(* Logix 5000 project; controller DSFW_0512_C_FCB_S1_SPN vendor 1 type 14 code 77 rev 20.12; software revision 20.06 *)

TASK MainTask (continuous, watchdog 500 ms) : General_Alarms_Config, Process_Control
TASK PID_Loops (periodic, rate 10 ms, priority 10, watchdog 500 ms) : Process_PID_Calculations

MODULES
   Controller : vendor 1 type 14 code 77 (CompactLogixL32EController 0, rev 20.12)
      LocalENB : 1769-L32E Ethernet Port (CompactLogixL32Ethernet 1, Ethernet 192.168.1.30, rev 20.11)
      Local : CompactBus (CompactVirtualAdapter 3, rev 20.11)
          : vendor 1 type 7 code 82 (Compact 1, rev 1.1, Input RPI 20 ms)
          : 1769-IF8 (Compact 3, rev 1.1, Output RPI 80 ms)
          : 1769-IR6 (Compact 4, rev 1.1, Input RPI 5 ms)
          : vendor 1 type 7 code 93 (Compact 2, rev 1.1, Output RPI 20 ms)
          : vendor 1 type 10 code 39 (Compact 5, rev 2.1, Output RPI 80 ms)
END_MODULES

VAR_GLOBAL   (* controller tags *)
   Alarms : DINT[3] := ([0] := 2);
   Alarms_Active : BOOL := 1;
   Batch_Mode_Enable : BOOL;
   Comp_Low_Pressure_Alarm_Setpoint : REAL := 12.0;
   Compressor_High_Pressure_Alarm_Setpoint : REAL := 300.0;
   Compressor_High_Pressure_Delay_Timer : TIMER := (PRE := 1000);
   Compressor_High_Superheat_Alarm_Delay : TIMER := (PRE := 600000);
   Compressor_High_Superheat_Alarm_Setpoint : REAL := 80.0;
   Compressor_Low_Pressure_Alarm_Setpoint : DINT := 120;
   Compressor_Low_Pressure_Delay_Timer : TIMER := (PRE := 60000);
   Compressor_Low_Subcooling_Alarm_Delay : TIMER := (PRE := 600000);
   Compressor_Low_Subcooling_Alarm_Setpoint : REAL := 4.0;
   Compressor_Low_Superheat_Alarm_Delay : TIMER := (PRE := 120000);
   Compressor_Low_Superheat_Alarm_Setpoint : REAL := 2.0;
   Compressor_OK_To_Run : BOOL;
   Compressor_Run_Proof_Delay : TIMER := (PRE := 5000);
   Compressor_Short_Cycle_Time_Remaining : REAL;
   Compressor_Short_Cycle_Timer : TIMER := (PRE := 60000);
   Compressor_Start_Delay : TIMER := (PRE := 10000);
   Compressor_Subcooling : REAL := 7.55085;
   Compressor_Superheat : REAL := 32.681896;
   Compresssor_Status : BOOL;
   Critical_Alarm : BOOL;
   DeltaV_Online : BOOL := 1;
   DeltaV_Status : DINT := 3;
   Display_Vessel_Select : BOOL;
   DV_IN_F8_50_99 : REAL[10] := ([0] := 11.0, [1] := 21.0, [2] := 21.0, [3] := 21.0); {produced}
   DV_IN_N7_100_199 : INT[10] := ([0] := 20, [1] := 4); {produced}
   DV_OUT_F8_0_49 : REAL[20] := ([0] := 21.3, [1] := 21.2, [2] := 10.7202635, [3] := -37.5, [4] := -37.5, [5] := -37.5, [8] := 109.89375, [9] := 180.79688, [10] := 79.402695, [11] := 8.548732, [13] := 74.6, [14] := 73.2, [15] := 84.7); {produced, access Read Only}
   DV_OUT_N7_0_99 : INT[20] := ([0] := 41, [1] := 16845, [2] := 3, [3] := 1, [4] := 2); {produced, access Read Only}
   EEV_101_Auto_Manual : BOOL;
   EEV_101_Manual_Output : REAL := 25.0;
   EEV_101_Output_Percent : REAL;
   EEV_101_Pressure_PIDE : PID_ENHANCED := (PV := 10.73405, PVEUMax := 103.0, PVEUMin := -7.3, SPProg := 125.0, SPOper := 125.0, SPHLimit := 103.0, SPLLimit := -7.3, RatioProg := 1.0, RatioOper := 1.0, RatioHLimit := 1.0, RatioLLimit := 1.0, CVEUMax := 10000.0, CVHLimit := 100.0, CVLLimit := 20.0, HandFB := 25.0, PGain := 10.0, IGain := 5.0, PVEDerivative := 1, ProgOverrideReq := 1, RTSTime := 1, CVLAlarm := 1, SP := 103.0, SPPercent := 100.0, SPHAlarm := 1, PVPercent := 16.35, E := 92.26595, EPercent := 83.65, InitPrimary := 1, WindupHOut := 1, WindupLOut := 1, Ratio := 1.0, Override := 1, DeltaT := 0.01, Status1 := 16#0000_0061, InstructFault := 1, SPProgInv := 1, SPOperInv := 1);
   EEV_101_Pressure_Setpoint : REAL := 125.0;
   EEV_101_Range_1_Max : REAL := 100.0;
   EEV_101_Range_1_Min : REAL := 20.0;
   EEV_101_Range_2_Max : REAL := 100.0;
   EEV_101_Range_2_Min : REAL := 20.0;
   EEV_101_Range_3_Max : REAL := 50.0;
   EEV_101_Range_3_Min : REAL := 10.0;
   EEV_101_Run_PIDE : BOOL;
   EEV_101_Run_Temp_PIDE : BOOL;
   EEV_101_Stop_PIDE : BOOL := 1;
   EEV_101_Superheat_PIDE : PID_ENHANCED := (PV := 21.081898, PVEUMax := 121.0, PVEUMin := -18.0, SPProg := 10.0, SPOper := 10.0, SPHLimit := 121.0, SPLLimit := -18.0, RatioProg := 1.0, RatioOper := 1.0, RatioHLimit := 1.0, RatioLLimit := 1.0, CVEUMax := 10000.0, CVHLimit := 100.0, CVLLimit := 20.0, HandFB := 25.0, ControlAction := 1, PGain := 10.0, IGain := 5.0, PVEDerivative := 1, ProgOverrideReq := 1, RTSTime := 1, CVLAlarm := 1, SP := 10.0, SPPercent := 20.143885, PVPercent := 28.116474, E := 11.081898, EPercent := 7.9725895, InitPrimary := 1, WindupHOut := 1, Ratio := 1.0, Override := 1, DeltaT := 0.01);
   EEV_101_Superheat_Setpoint : REAL := 10.0;
   EEV_101_Temperature_PIDE : PID_ENHANCED := (PV := 21.3, PVEUMax := 121.0, PVEUMin := -18.0, SPProg := 11.0, SPOper := 11.0, SPCascade := 11.0, SPHLimit := 121.0, SPLLimit := -18.0, RatioProg := 1.0, RatioOper := 1.0, RatioHLimit := 1.0, RatioLLimit := 1.0, CVEUMax := 10000.0, CVHLimit := 100.0, CVLLimit := 20.0, HandFB := 25.0, ControlAction := 1, PGain := 10.0, IGain := 5.0, PVEDerivative := 1, AllowCasRat := 1, ProgOverrideReq := 1, RTSTime := 1, CVLAlarm := 1, SP := 11.0, SPPercent := 20.86331, PVPercent := 28.27338, E := 10.299999, EPercent := 7.4100704, InitPrimary := 1, WindupHOut := 1, Ratio := 1.0, Override := 1, DeltaT := 0.01);
   EEV_102_Auto_Manual : BOOL;
   EEV_102_Manual_Output : REAL := 12.0;
   EEV_102_Output_Percent : REAL;
   EEV_102_PIDE : PID_ENHANCED := (PV := 32.681896, PVEUMax := 121.0, PVEUMin := -18.0, SPProg := 50.0, SPOper := 50.0, SPHLimit := 121.0, SPLLimit := -18.0, RatioProg := 1.0, RatioOper := 1.0, RatioHLimit := 1.0, RatioLLimit := 1.0, CVEUMax := 10000.0, CVHLimit := 100.0, HandFB := 12.0, ControlAction := 1, PGain := 0.3, IGain := 0.1, PVEDerivative := 1, ProgOverrideReq := 1, RTSTime := 1, SP := 50.0, SPPercent := 48.920864, PVPercent := 36.461796, E := -17.318104, EPercent := -12.459068, InitPrimary := 1, Ratio := 1.0, Override := 1, DeltaT := 0.01);
   EEV_102_SH_Setpoint : REAL := 50.0;
   EEV_102_Stop_PIDE : BOOL := 1;
   Enable_Batch : BOOL := 1;
   Evaporator_Low_Flow_Delay_Timer : TIMER;
   Evaporator_Low_Flow_Setpoint : REAL;
   Evaporator_Low_Superheat_Alarm_Delay : TIMER := (PRE := 120);
   Evaporator_Low_Superheat_Alarm_Setpoint : REAL;
   Evaporator_Superheat : REAL := 21.081898;
   Glycol_Skid_Run : BOOL;
   Glycol_Skid_Status : BOOL;
   Heater_Start_Delay : TIMER := (PRE := 5000);
   Heaters_OK_To_Run : BOOL;
   HMI_Compressor_High_Superheat_Delay : REAL := 600.0;
   HMI_Compressor_Low_Pressure_Delay : REAL := 60.0;
   HMI_Compressor_Low_Subcooling_Delay : REAL := 600.0;
   HMI_Compressor_Low_Superheat_Delay : REAL := 120.0;
   HMI_Evaporator_Low_Superheat_Delay : REAL := 120.0;
   HMI_Pump_High_Pressure_Delay : REAL;
   HMI_Pump_Low_Pressure_Delay : REAL := 20.0;
   HMI_Remote_Enable : BOOL := 1;
   HMI_Tank_High_Pressure_Delay : REAL := 5.0;
   HMI_Tank_Low_Level_Delay : REAL := 10.0;
   Jacket_High_High_Temperature_Setpoint : REAL := 110.0;
   Jacket_High_Temperature_Setpoint : REAL := 110.0;
   Jacket_Low_Low_Temperature_Setpoint : REAL := -20.0;
   Jacket_Low_Temperature_Setpoint : REAL := -20.0;
   Large_Batch_Derivative : REAL;
   Large_Batch_Integral : REAL := 0.9;
   Large_Batch_Proportional : REAL := 15.0;
   Large_Batch_Selected : BOOL;
   LSH_101_Status : BOOL := 1;
   LSL_101_Status : BOOL := 1;
   LSL_102_Status : BOOL := 1;
   Medium_Batch_Derivative : REAL;
   Medium_Batch_Integral : REAL := 0.9;
   Medium_Batch_Proportional : REAL := 15.0;
   Medium_Batch_Selected : BOOL;
   Phase_Monitor_Delay : TIMER := (PRE := 5000);
   Process_Pump_Flow_Rate : REAL := -45.73986;
   Process_Pump_Low_Flow_Alarm_Setpoint : DINT;
   PT_101_Offset : REAL;
   PT_101_Reactor_Supply_Pressure : REAL := 10.713368;
   PT_101_Sensor_Alarm_Delay : TIMER := (PRE := 5000);
   PT_102_Compressor_Suction_Pressure : REAL := 109.89375;
   PT_102_Offset : REAL;
   PT_102_Sensor_Alarm_Delay : TIMER := (PRE := 5000);
   PT_103_Compressor_Discharge_Pressure : REAL := 180.79688;
   PT_103_Offset : REAL;
   PT_103_Sensor_Alarm_Delay : TIMER := (PRE := 5000);
   PT_104_Evaporator_Suction_Pressure : REAL := 109.89375;
   PT_104_Offset : REAL;
   PT_104_Sensor_Alarm_Delay : TIMER := (PRE := 5000);
   PT_105_Offset : REAL;
   PT_105_Sensor_Alarm_Delay : TIMER := (PRE := 5000);
   PT_105_Tank_Blanket_Pressure : REAL := 8.562519;
   Pump_High_Pressure_Delay : TIMER;
   Pump_High_Pressure_Setpoint : REAL := 100.0;
   Pump_Low_Flow_Delay_Timer : TIMER;
   Pump_Low_Pressure_Delay : TIMER := (PRE := 20000);
   Pump_Low_Pressure_Setpoint : REAL := 5.0;
   Pump_OK_To_Run : BOOL;
   Pump_Start_Delay : TIMER := (PRE := 5000);
   Pump_Status : BOOL;
   Reaactor_Batch_PIDE : PID_ENHANCED := (PV := -37.5, PVEUMax := 100.0, PVEUMin := -15.0, SPProg := 11.0, SPOper := -15.0, SPHLimit := 100.0, SPLLimit := -15.0, RatioProg := 1.0, RatioOper := 1.0, RatioHLimit := 1.0, RatioLLimit := 1.0, CVInitReq := 1, CVInitValue := 11.0, CVEUMax := -32.5, CVEUMin := -5.0, CVHLimit := 100.0, PGain := 15.0, IGain := 0.9, PVEDerivative := 1, DSmoothing := 1, PVTracking := 1, ManualAfterInit := 1, ProgOverrideReq := 1, RTSTime := 1, CVEU := 11.0, CVInitializing := 1, CVLAlarm := 1, SP := -15.0, SPLAlarm := 1, PVPercent := -19.565218, E := 22.5, EPercent := 19.565218, InitPrimary := 1, Ratio := 1.0, Override := 1, DeltaT := 0.01);
   Reactor_Batch_CV_as_SP : REAL := 11.0;
   Reactor_Batch_PID_Start : BOOL;
   Reactor_Batch_PID_Start_Delay : TIMER := (PRE := 5000);
   Reactor_Batch_PID_Start_ONS : BOOL;
   Reactor_Batch_PID_Stop : BOOL := 1;
   Reactor_Batch_PV : REAL := -37.5;
   Reactor_Batch_SP_High : REAL := -32.5;
   Reactor_Batch_SP_Low : REAL := -42.5;
   Read_PLC_Clock : DINT[7] := ([0] := 1999, [1] := 12, [2] := 29, [3] := 18, [4] := 28, [5] := 41, [6] := 799818);
   Remote_Enable : BOOL := 1;
   Remote_Start : BOOL;
   Reset_Alarms : BOOL;
   Reset_Defaults : BOOL;
   SCR_101_Auto_Manual : BOOL;
   SCR_101_Manual_Output : REAL;
   SCR_101_Output_Percent : REAL;
   SCR_101_PIDE : PID_ENHANCED := (PV := 21.3, PVEUMax := 121.0, PVEUMin := -18.0, SPProg := 11.0, SPOper := 21.3, SPCascade := 11.0, SPHLimit := 121.0, SPLLimit := -18.0, RatioProg := 1.0, RatioOper := 1.0, RatioHLimit := 1.0, RatioLLimit := 1.0, CVEUMax := 10000.0, CVHLimit := 100.0, PGain := 50.0, IGain := 5.0, PVEDerivative := 1, PVTracking := 1, AllowCasRat := 1, ProgOverrideReq := 1, RTSTime := 1, SP := 21.3, SPPercent := 28.27338, PVPercent := 28.27338, InitPrimary := 1, Ratio := 1.0, Override := 1, DeltaT := 0.01);
   SCR_101_Run_PIDE : BOOL;
   SCR_101_Stop_PIDE : BOOL := 1;
   Select_Large_Batch : BOOL;
   Select_Medium_Batch : BOOL;
   Select_Small_Batch : BOOL;
   Select_Vessel_1 : BOOL;
   Select_Vessel_2 : BOOL;
   Select_Vessel_3 : BOOL;
   Show_Local : BOOL;
   SIC_101_Auto_Manual : BOOL;
   SIC_101_Manual_Output : REAL := 100.0;
   SIC_101_Output_Percent : REAL;
   SIC_101_PIDE : PID_ENHANCED := (PV := 10.740945, PVEUMax := 103.0, PVEUMin := -7.3, SPProg := 50.0, SPOper := 50.0, SPHLimit := 103.0, SPLLimit := -7.3, RatioProg := 1.0, RatioOper := 1.0, RatioHLimit := 1.0, RatioLLimit := 1.0, CVEUMax := 10000.0, CVHLimit := 100.0, HandFB := 100.0, IGain := 10.0, PVEDerivative := 1, ProgOverrideReq := 1, RTSTime := 1, SP := 50.0, SPPercent := 51.949226, PVPercent := 16.35625, E := 39.259056, EPercent := 35.592976, InitPrimary := 1, Ratio := 1.0, Override := 1, DeltaT := 0.01);
   SIC_101_Pressure_Setpoint : REAL := 50.0;
   SIC_101_Run_PIDE : BOOL;
   SIC_101_Stop_PIDE : BOOL := 1;
   Small_Batch_Derivative : REAL;
   Small_Batch_Integral : REAL := 0.9;
   Small_Batch_Proportional : REAL := 15.0;
   Small_Batch_Selected : BOOL;
   SP_Add_Max : REAL := 5.0;
   SP_Add_Min : REAL := 50.0;
   Startup_Delay : TIMER := (PRE := 250, ACC := 250, EN := 1, DN := 1);
   System_Start : BOOL := 1;
   Tank_High_Pressure_Delay : TIMER := (PRE := 5000);
   Tank_High_Pressure_Setpoint : REAL := 15.0;
   Tank_Low_Level_Delay : TIMER := (PRE := 10000);
   TCV_101_Auto_Manual : BOOL;
   TCV_101_Define_Range_1_Max : REAL := -5.0;
   TCV_101_Define_Range_1_Min : REAL := -30.0;
   TCV_101_Define_Range_2_Max : REAL := 50.0;
   TCV_101_Define_Range_2_Min : REAL := -4.9;
   TCV_101_Define_Range_3_Max : REAL := 130.0;
   TCV_101_Define_Range_3_Min : REAL := 50.1;
   TCV_101_Manual_Output : REAL;
   TCV_101_Output_Percent : REAL;
   TCV_101_PIDE : PID_ENHANCED := (PV := 21.3, PVEUMax := 121.0, PVEUMin := -18.0, SPProg := 11.0, SPOper := 11.0, SPCascade := 11.0, SPHLimit := 121.0, SPLLimit := -18.0, RatioProg := 1.0, RatioOper := 1.0, RatioHLimit := 1.0, RatioLLimit := 1.0, CVEUMax := 10000.0, CVHLimit := 50.0, CVLLimit := 15.0, PGain := 10.0, IGain := 5.0, PVEDerivative := 1, AllowCasRat := 1, ProgOverrideReq := 1, RTSTime := 1, CVLAlarm := 1, SP := 11.0, SPPercent := 20.86331, PVPercent := 28.27338, E := -10.299999, EPercent := -7.4100704, InitPrimary := 1, WindupLOut := 1, Ratio := 1.0, Override := 1, DeltaT := 0.01);
   TCV_101_Range_1_Max : REAL := 50.0;
   TCV_101_Range_1_Min : REAL := 15.0;
   TCV_101_Range_2_Max : REAL := 50.0;
   TCV_101_Range_2_Min : REAL := 15.0;
   TCV_101_Range_3_Max : REAL := 50.0;
   TCV_101_Range_3_Min : REAL := 5.0;
   TCV_101_Run_PIDE : BOOL;
   TCV_101_Stop_PIDE : BOOL := 1;
   TE_101_Liquid_Line_Temperature : REAL := 74.6;
   TE_101_Offset : REAL;
   TE_102_Evaporator_Suction_Temperature : REAL := 73.1;
   TE_102_Offset : REAL;
   TE_103_Compressor_Suction_Temperature : REAL := 84.6;
   TE_103_Offset : REAL;
   TE_104_Offset : REAL;
   TE_104_Reactor_Return_Temperature : REAL := 21.2;
   TE_105_Offset : REAL;
   TE_105_Reactor_Supply_Temperature : REAL := 21.3;
   Temperature_Setpoint : REAL := 11.0;
   Test_Analog : REAL := 4000.0;
   Test_Bit : BOOL[32] := ([0] := 1, [1] := 1);
   TIT_101_Offset : REAL;
   TIT_101_Sensor_Alarm_Delay : TIMER := (PRE := 5000);
   TIT_101_Vessel_Temperature : REAL := -37.5;
   TIT_201_Offset : REAL;
   TIT_201_Sensor_Alarm_Delay : TIMER;
   TIT_201_Vessel_Temperature : REAL := -37.5;
   TIT_301_Offset : REAL;
   TIT_301_Sensor_Alarm_Delay : TIMER;
   TIT_301_Vessel_Temperature : REAL := -37.5;
   Vessel_1_Scale_Max : REAL := 120.0;
   Vessel_1_Scale_Min : REAL := -30.0;
   Vessel_1_Selected : BOOL;
   Vessel_2_Scale_Max : REAL := 120.0;
   Vessel_2_Scale_Min : REAL := -30.0;
   Vessel_2_Selected : BOOL;
   Vessel_3_Scale_Max : REAL := 120.0;
   Vessel_3_Scale_Min : REAL := -30.0;
   Vessel_3_Selected : BOOL;
   Vessel_High_High_Temperature_Setpoint : REAL := 110.0;
   Vessel_High_Temperature_Setpoint : REAL := 110.0;
   Vessel_Low_Low_Temperature_Setpoint : REAL := -20.0;
   Vessel_Low_Temperature_Setpoint : REAL := -20.0;
   Warning_Alarms : BOOL := 1;
END_VAR

PROGRAM General_Alarms_Config   (* main routine MainRoutine *)

ROUTINE DV_Communications   (* ladder *)
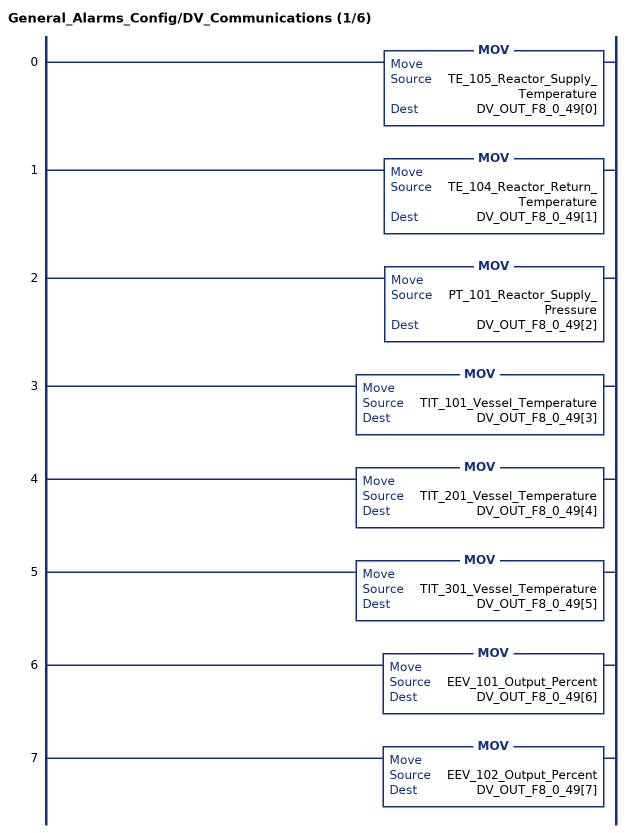
   0: MOV(TE_105_Reactor_Supply_Temperature,DV_OUT_F8_0_49[0]);
   1: MOV(TE_104_Reactor_Return_Temperature,DV_OUT_F8_0_49[1]);
   2: MOV(PT_101_Reactor_Supply_Pressure,DV_OUT_F8_0_49[2]);
   3: MOV(TIT_101_Vessel_Temperature,DV_OUT_F8_0_49[3]);
   4: MOV(TIT_201_Vessel_Temperature,DV_OUT_F8_0_49[4]);
   5: MOV(TIT_301_Vessel_Temperature,DV_OUT_F8_0_49[5]);
   6: MOV(EEV_101_Output_Percent,DV_OUT_F8_0_49[6]);
   7: MOV(EEV_102_Output_Percent,DV_OUT_F8_0_49[7]);
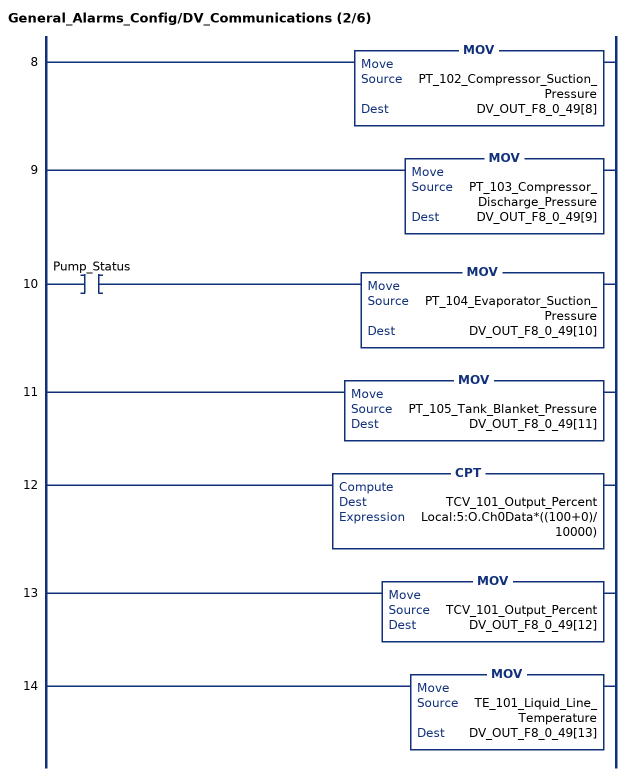
   8: MOV(PT_102_Compressor_Suction_Pressure,DV_OUT_F8_0_49[8]);
   9: MOV(PT_103_Compressor_Discharge_Pressure,DV_OUT_F8_0_49[9]);
   10: XIC(Pump_Status)MOV(PT_104_Evaporator_Suction_Pressure,DV_OUT_F8_0_49[10]);
   11: MOV(PT_105_Tank_Blanket_Pressure,DV_OUT_F8_0_49[11]);
   12: CPT(TCV_101_Output_Percent,Local:5:O.Ch0Data*((100+0)/10000));
   13: MOV(TCV_101_Output_Percent,DV_OUT_F8_0_49[12]);
   14: MOV(TE_101_Liquid_Line_Temperature,DV_OUT_F8_0_49[13]);
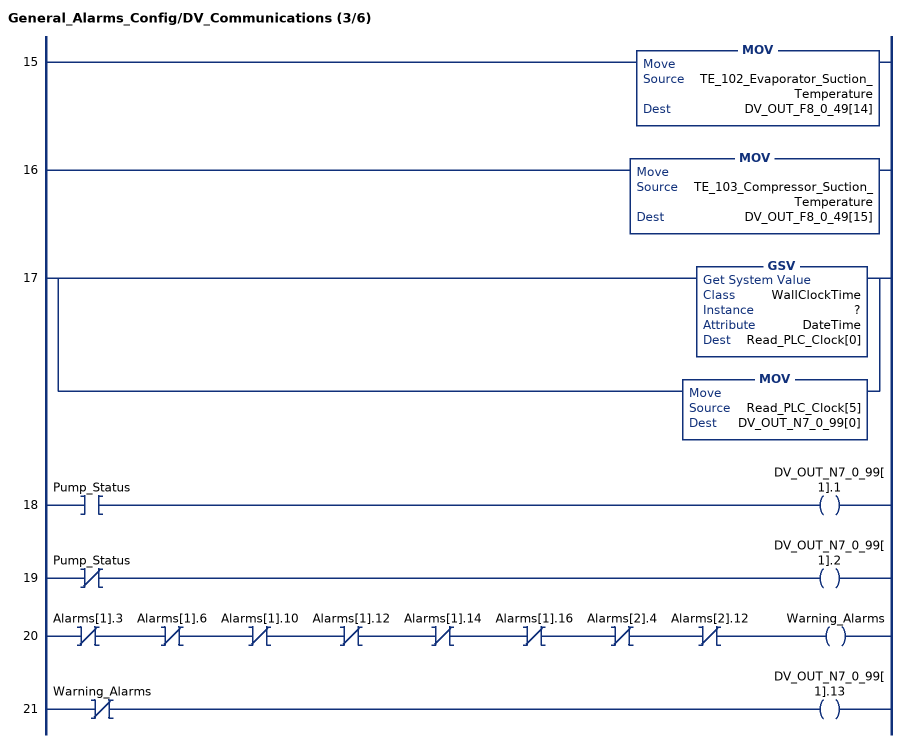
   15: MOV(TE_102_Evaporator_Suction_Temperature,DV_OUT_F8_0_49[14]);
   16: MOV(TE_103_Compressor_Suction_Temperature,DV_OUT_F8_0_49[15]);
   17: [GSV(WallClockTime,?,DateTime,Read_PLC_Clock[0]) ,MOV(Read_PLC_Clock[5],DV_OUT_N7_0_99[0]) ];
   18: XIC(Pump_Status)OTE(DV_OUT_N7_0_99[1].1);
   19: XIO(Pump_Status)OTE(DV_OUT_N7_0_99[1].2);
   20: XIO(Alarms[1].3)XIO(Alarms[1].6)XIO(Alarms[1].10)XIO(Alarms[1].12)XIO(Alarms[1].14)XIO(Alarms[1].16)XIO(Alarms[2].4)XIO(Alarms[2].12)OTE(Warning_Alarms);
   21: XIO(Warning_Alarms)OTE(DV_OUT_N7_0_99[1].13);
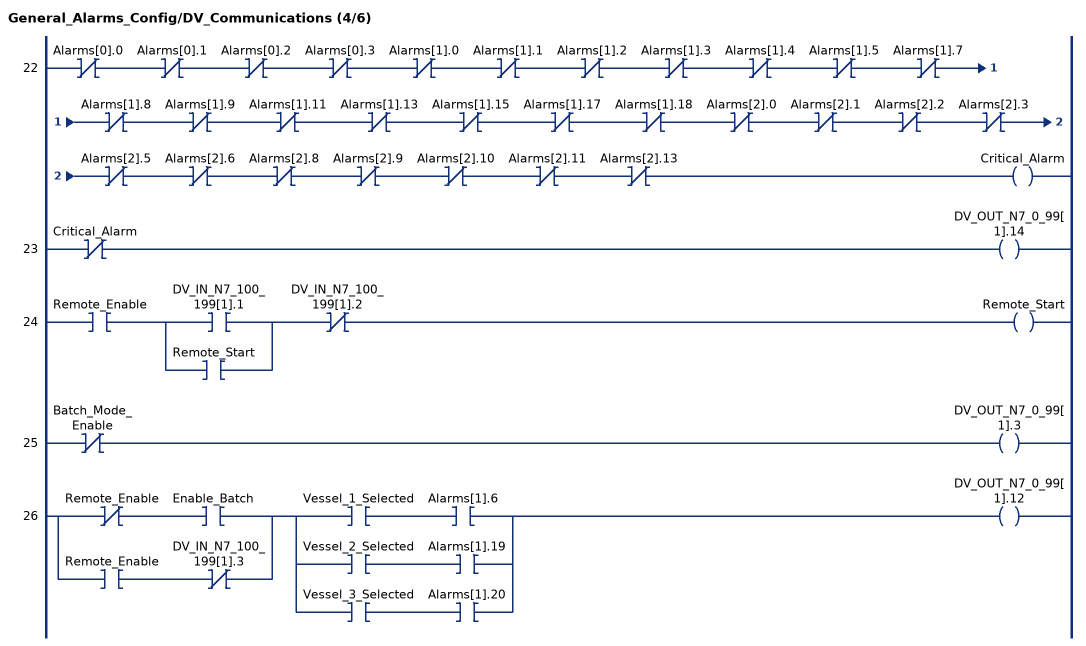
   22: XIO(Alarms[0].0)XIO(Alarms[0].1)XIO(Alarms[0].2)XIO(Alarms[0].3)XIO(Alarms[1].0)XIO(Alarms[1].1)XIO(Alarms[1].2)XIO(Alarms[1].3)XIO(Alarms[1].4)XIO(Alarms[1].5)XIO(Alarms[1].7)XIO(Alarms[1].8)XIO(Alarms[1].9)XIO(Alarms[1].11)XIO(Alarms[1].13)XIO(Alarms[1].15)XIO(Alarms[1].17)XIO(Alarms[1].18)XIO(Alarms[2].0)XIO(Alarms[2].1)XIO(Alarms[2].2)XIO(Alarms[2].3)XIO(Alarms[2].5)XIO(Alarms[2].6)XIO(Alarms[2].8)XIO(Alarms[2].9)XIO(Alarms[2].10)XIO(Alarms[2].11)XIO(Alarms[2].13)OTE(Critical_Alarm);
   23: XIO(Critical_Alarm)OTE(DV_OUT_N7_0_99[1].14);
   24: XIC(Remote_Enable)[XIC(DV_IN_N7_100_199[1].1) ,XIC(Remote_Start) ]XIO(DV_IN_N7_100_199[1].2)OTE(Remote_Start);
   25: XIO(Batch_Mode_Enable)OTE(DV_OUT_N7_0_99[1].3);
   26: [XIO(Remote_Enable) XIC(Enable_Batch) ,XIC(Remote_Enable) XIO(DV_IN_N7_100_199[1].3) ][XIC(Vessel_1_Selected) XIC(Alarms[1].6) ,XIC(Vessel_2_Selected) XIC(Alarms[1].19) ,XIC(Vessel_3_Selected) XIC(Alarms[1].20) ]OTE(DV_OUT_N7_0_99[1].12);
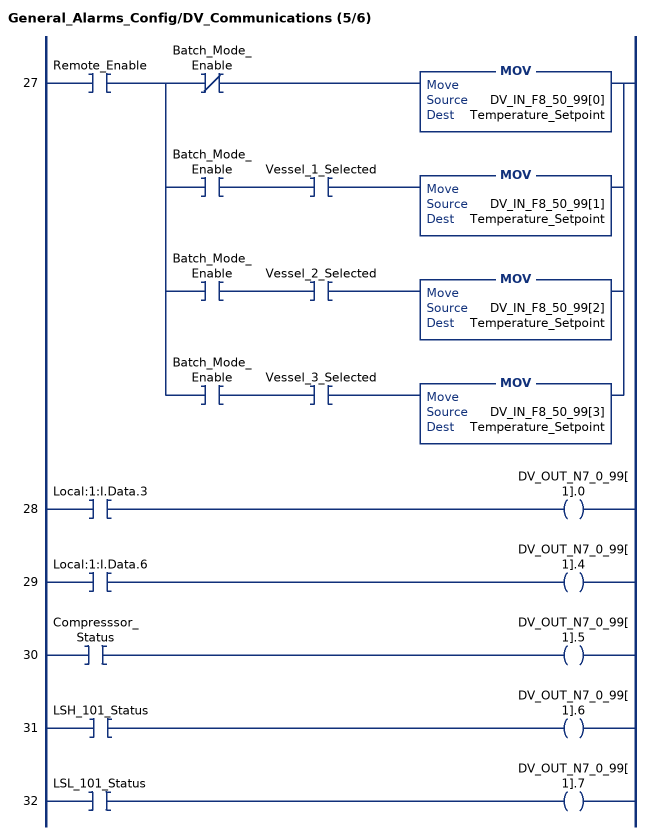
   27: XIC(Remote_Enable)[XIO(Batch_Mode_Enable) MOV(DV_IN_F8_50_99[0],Temperature_Setpoint) ,XIC(Batch_Mode_Enable) XIC(Vessel_1_Selected) MOV(DV_IN_F8_50_99[1],Temperature_Setpoint) ,XIC(Batch_Mode_Enable) XIC(Vessel_2_Selected) MOV(DV_IN_F8_50_99[2],Temperature_Setpoint) ,XIC(Batch_Mode_Enable) XIC(Vessel_3_Selected) MOV(DV_IN_F8_50_99[3],Temperature_Setpoint) ];
   28: XIC(Local:1:I.Data.3)OTE(DV_OUT_N7_0_99[1].0);
   29: XIC(Local:1:I.Data.6)OTE(DV_OUT_N7_0_99[1].4);
   30: XIC(Compresssor_Status)OTE(DV_OUT_N7_0_99[1].5);
   31: XIC(LSH_101_Status)OTE(DV_OUT_N7_0_99[1].6);
   32: XIC(LSL_101_Status)OTE(DV_OUT_N7_0_99[1].7);
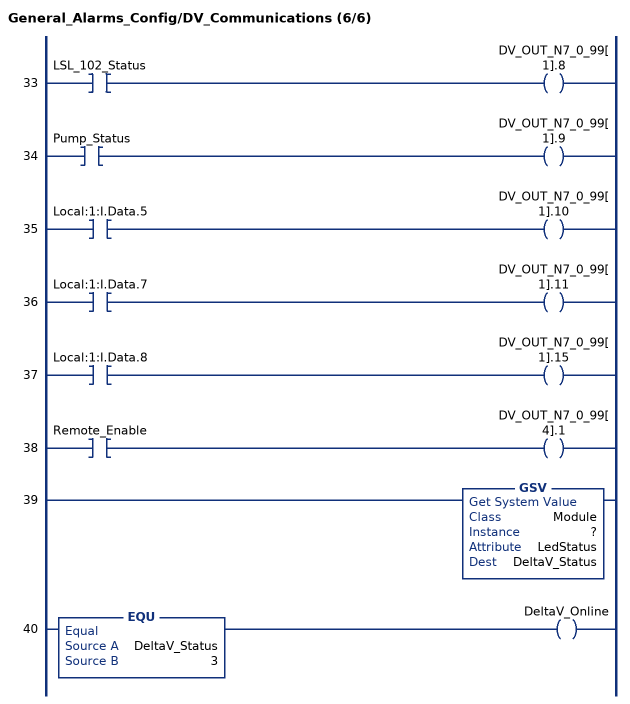
   33: XIC(LSL_102_Status)OTE(DV_OUT_N7_0_99[1].8);
   34: XIC(Pump_Status)OTE(DV_OUT_N7_0_99[1].9);
   35: XIC(Local:1:I.Data.5)OTE(DV_OUT_N7_0_99[1].10);
   36: XIC(Local:1:I.Data.7)OTE(DV_OUT_N7_0_99[1].11);
   37: XIC(Local:1:I.Data.8)OTE(DV_OUT_N7_0_99[1].15);
   38: XIC(Remote_Enable)OTE(DV_OUT_N7_0_99[4].1);
   39: GSV(Module,?,LedStatus,DeltaV_Status);
   40: EQU(DeltaV_Status,3)OTE(DeltaV_Online);
END_ROUTINE

ROUTINE HMI_Writes   (* ladder *)
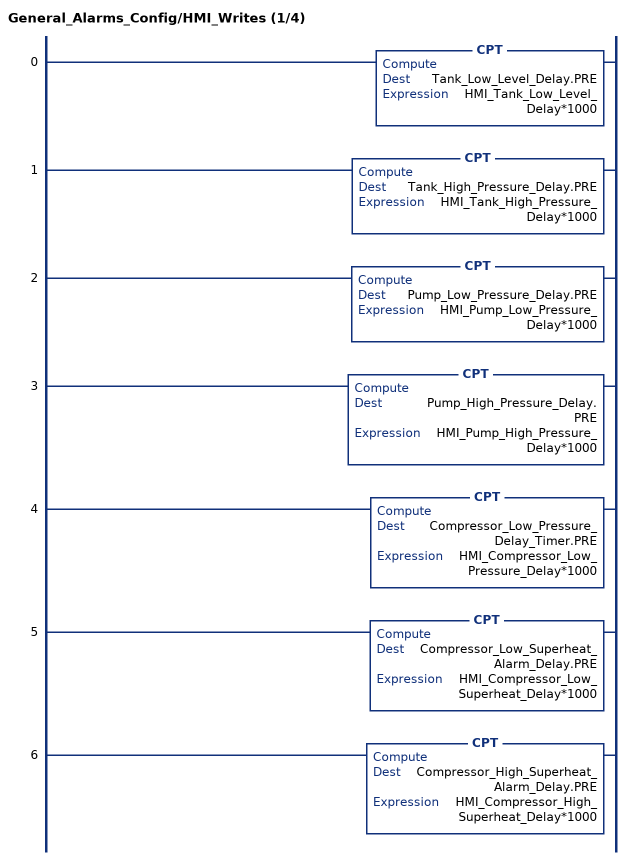
   0: CPT(Tank_Low_Level_Delay.PRE,HMI_Tank_Low_Level_Delay*1000);
   1: CPT(Tank_High_Pressure_Delay.PRE,HMI_Tank_High_Pressure_Delay*1000);
   2: CPT(Pump_Low_Pressure_Delay.PRE,HMI_Pump_Low_Pressure_Delay*1000);
   3: CPT(Pump_High_Pressure_Delay.PRE,HMI_Pump_High_Pressure_Delay*1000);
   4: CPT(Compressor_Low_Pressure_Delay_Timer.PRE,HMI_Compressor_Low_Pressure_Delay*1000);
   5: CPT(Compressor_Low_Superheat_Alarm_Delay.PRE,HMI_Compressor_Low_Superheat_Delay*1000);
   6: CPT(Compressor_High_Superheat_Alarm_Delay.PRE,HMI_Compressor_High_Superheat_Delay*1000);
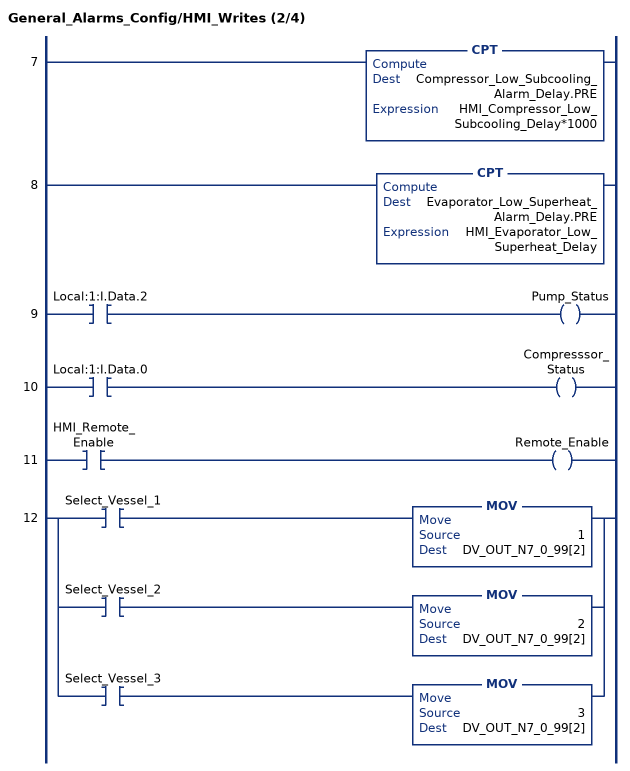
   7: CPT(Compressor_Low_Subcooling_Alarm_Delay.PRE,HMI_Compressor_Low_Subcooling_Delay*1000);
   8: CPT(Evaporator_Low_Superheat_Alarm_Delay.PRE,HMI_Evaporator_Low_Superheat_Delay);
   9: XIC(Local:1:I.Data.2)OTE(Pump_Status);
   10: XIC(Local:1:I.Data.0)OTE(Compresssor_Status);
   11: XIC(HMI_Remote_Enable)OTE(Remote_Enable);
   12: [XIC(Select_Vessel_1) MOV(1,DV_OUT_N7_0_99[2]) ,XIC(Select_Vessel_2) MOV(2,DV_OUT_N7_0_99[2]) ,XIC(Select_Vessel_3) MOV(3,DV_OUT_N7_0_99[2]) ];
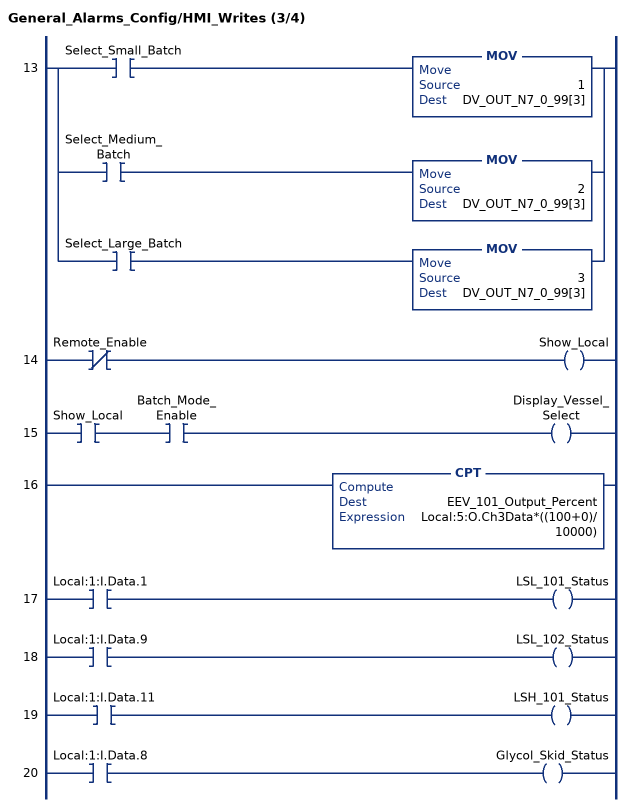
   13: [XIC(Select_Small_Batch) MOV(1,DV_OUT_N7_0_99[3]) ,XIC(Select_Medium_Batch) MOV(2,DV_OUT_N7_0_99[3]) ,XIC(Select_Large_Batch) MOV(3,DV_OUT_N7_0_99[3]) ];
   14: XIO(Remote_Enable)OTE(Show_Local);
   15: XIC(Show_Local)XIC(Batch_Mode_Enable)OTE(Display_Vessel_Select);
   16: CPT(EEV_101_Output_Percent,Local:5:O.Ch3Data*((100+0)/10000));
   17: XIC(Local:1:I.Data.1)OTE(LSL_101_Status);
   18: XIC(Local:1:I.Data.9)OTE(LSL_102_Status);
   19: XIC(Local:1:I.Data.11)OTE(LSH_101_Status);
   20: XIC(Local:1:I.Data.8)OTE(Glycol_Skid_Status);
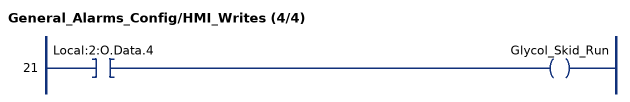
   21: XIC(Local:2:O.Data.4)OTE(Glycol_Skid_Run);
END_ROUTINE

ROUTINE MainRoutine   (* ladder *)
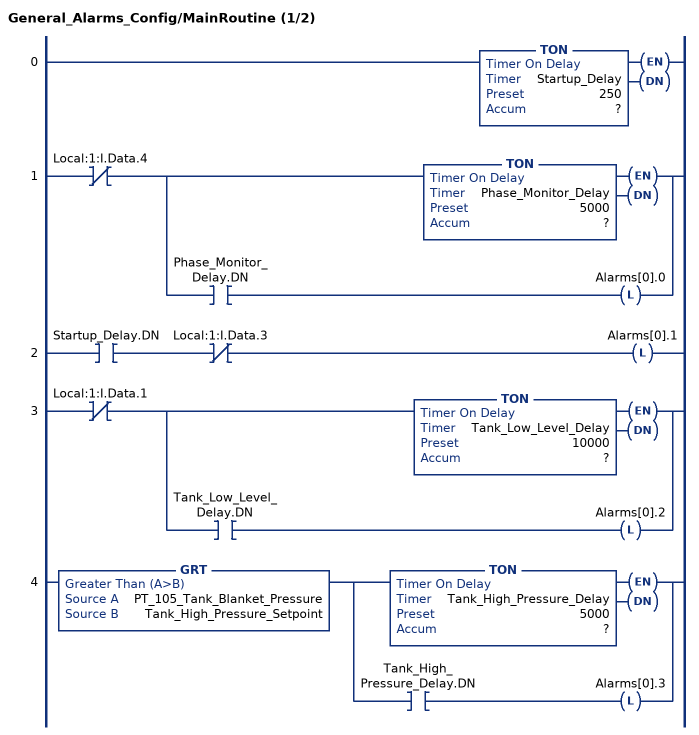
   0: TON(Startup_Delay,?,?);
   1: XIO(Local:1:I.Data.4)[TON(Phase_Monitor_Delay,?,?) ,XIC(Phase_Monitor_Delay.DN) OTL(Alarms[0].0) ];
   2: XIC(Startup_Delay.DN)XIO(Local:1:I.Data.3)OTL(Alarms[0].1);
   3: XIO(Local:1:I.Data.1)[TON(Tank_Low_Level_Delay,?,?) ,XIC(Tank_Low_Level_Delay.DN) OTL(Alarms[0].2) ];
   4: GRT(PT_105_Tank_Blanket_Pressure,Tank_High_Pressure_Setpoint)[TON(Tank_High_Pressure_Delay,?,?) ,XIC(Tank_High_Pressure_Delay.DN) OTL(Alarms[0].3) ];
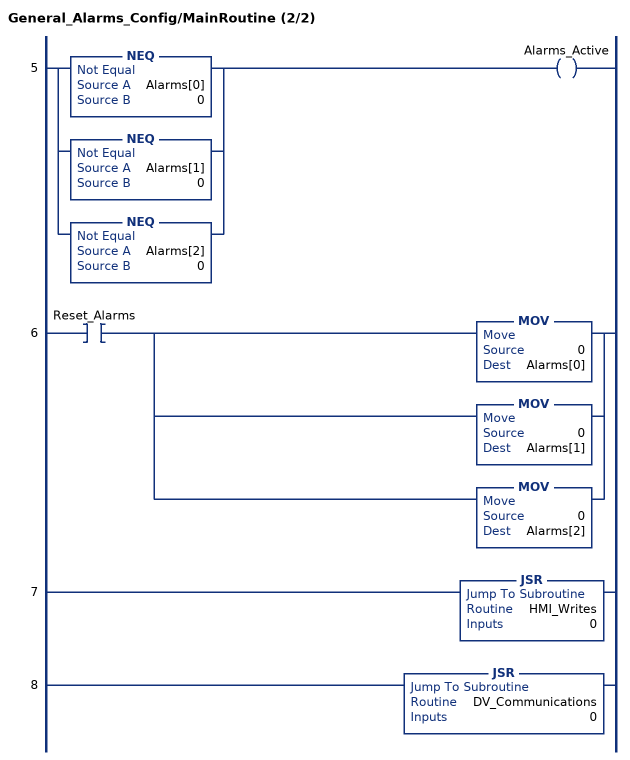
   5: [NEQ(Alarms[0],0) ,NEQ(Alarms[1],0) ,NEQ(Alarms[2],0) ]OTE(Alarms_Active);
   6: XIC(Reset_Alarms)[MOV(0,Alarms[0]) ,MOV(0,Alarms[1]) ,MOV(0,Alarms[2]) ];
   7: JSR(HMI_Writes,0);
   8: JSR(DV_Communications,0);
END_ROUTINE
END_PROGRAM

PROGRAM Process_Control   (* main routine Config *)

ROUTINE Alarms   (* ladder *)
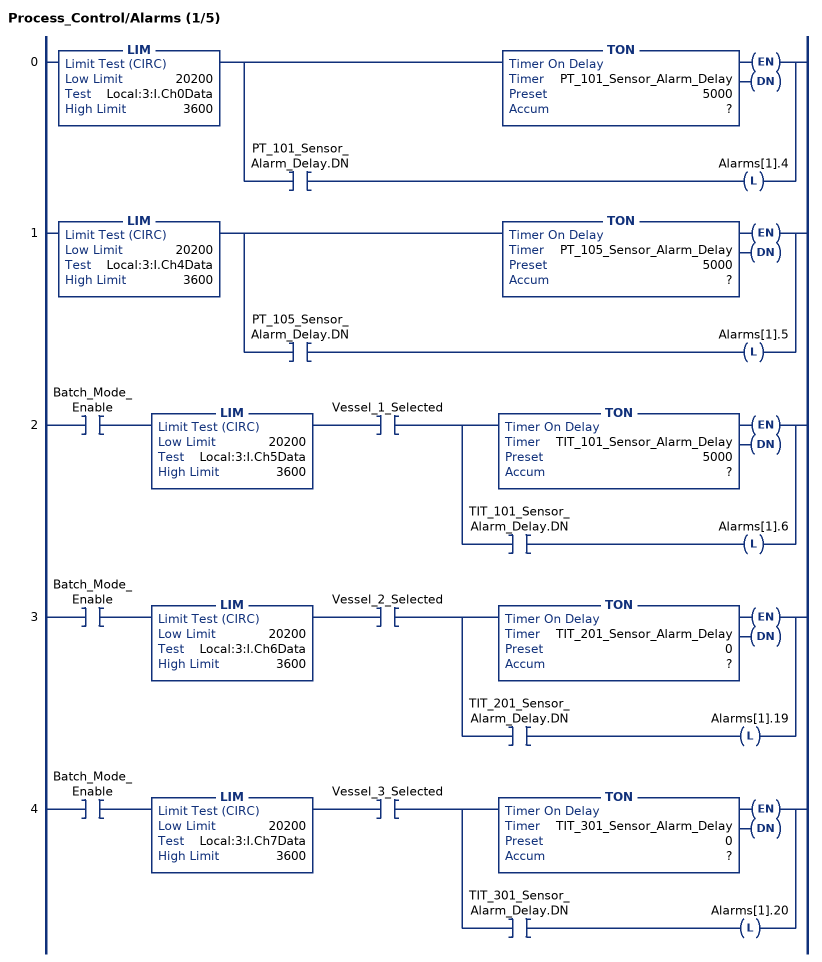
   0: LIM(20200,Local:3:I.Ch0Data,3600)[TON(PT_101_Sensor_Alarm_Delay,?,?) ,XIC(PT_101_Sensor_Alarm_Delay.DN) OTL(Alarms[1].4) ];
   1: LIM(20200,Local:3:I.Ch4Data,3600)[TON(PT_105_Sensor_Alarm_Delay,?,?) ,XIC(PT_105_Sensor_Alarm_Delay.DN) OTL(Alarms[1].5) ];
   2: XIC(Batch_Mode_Enable)LIM(20200,Local:3:I.Ch5Data,3600)XIC(Vessel_1_Selected)[TON(TIT_101_Sensor_Alarm_Delay,?,?) ,XIC(TIT_101_Sensor_Alarm_Delay.DN) OTL(Alarms[1].6) ];
   3: XIC(Batch_Mode_Enable)LIM(20200,Local:3:I.Ch6Data,3600)XIC(Vessel_2_Selected)[TON(TIT_201_Sensor_Alarm_Delay,?,?) ,XIC(TIT_201_Sensor_Alarm_Delay.DN) OTL(Alarms[1].19) ];
   4: XIC(Batch_Mode_Enable)LIM(20200,Local:3:I.Ch7Data,3600)XIC(Vessel_3_Selected)[TON(TIT_301_Sensor_Alarm_Delay,?,?) ,XIC(TIT_301_Sensor_Alarm_Delay.DN) OTL(Alarms[1].20) ];
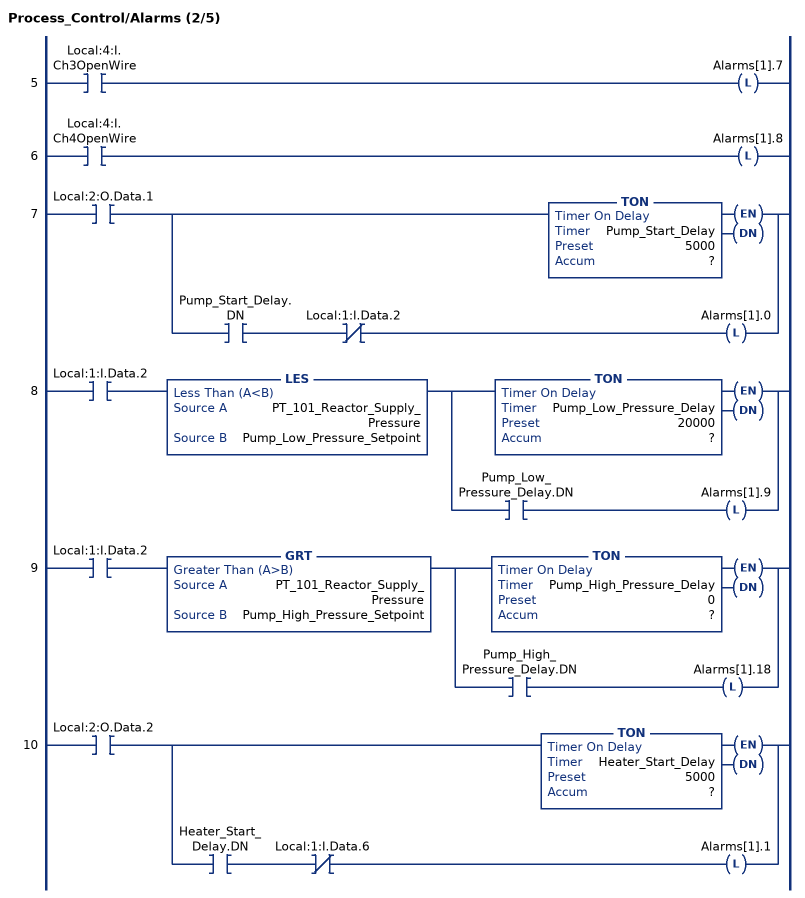
   5: XIC(Local:4:I.Ch3OpenWire)OTL(Alarms[1].7);
   6: XIC(Local:4:I.Ch4OpenWire)OTL(Alarms[1].8);
   7: XIC(Local:2:O.Data.1)[TON(Pump_Start_Delay,?,?) ,XIC(Pump_Start_Delay.DN) XIO(Local:1:I.Data.2) OTL(Alarms[1].0) ];
   8: XIC(Local:1:I.Data.2)LES(PT_101_Reactor_Supply_Pressure,Pump_Low_Pressure_Setpoint)[TON(Pump_Low_Pressure_Delay,?,?) ,XIC(Pump_Low_Pressure_Delay.DN) OTL(Alarms[1].9) ];
   9: XIC(Local:1:I.Data.2)GRT(PT_101_Reactor_Supply_Pressure,Pump_High_Pressure_Setpoint)[TON(Pump_High_Pressure_Delay,?,?) ,XIC(Pump_High_Pressure_Delay.DN) OTL(Alarms[1].18) ];
   10: XIC(Local:2:O.Data.2)[TON(Heater_Start_Delay,?,?) ,XIC(Heater_Start_Delay.DN) XIO(Local:1:I.Data.6) OTL(Alarms[1].1) ];
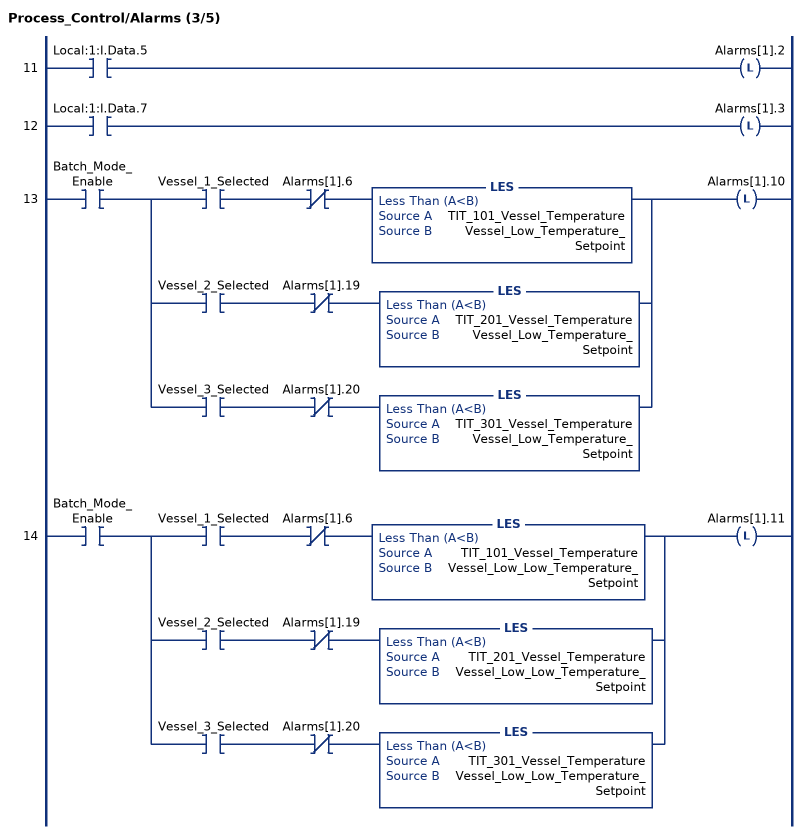
   11: XIC(Local:1:I.Data.5)OTL(Alarms[1].2);
   12: XIC(Local:1:I.Data.7)OTL(Alarms[1].3);
   13: XIC(Batch_Mode_Enable)[XIC(Vessel_1_Selected) XIO(Alarms[1].6) LES(TIT_101_Vessel_Temperature,Vessel_Low_Temperature_Setpoint) ,XIC(Vessel_2_Selected) XIO(Alarms[1].19) LES(TIT_201_Vessel_Temperature,Vessel_Low_Temperature_Setpoint) ,XIC(Vessel_3_Selected) XIO(Alarms[1].20) LES(TIT_301_Vessel_Temperature,Vessel_Low_Temperature_Setpoint) ]OTL(Alarms[1].10);
   14: XIC(Batch_Mode_Enable)[XIC(Vessel_1_Selected) XIO(Alarms[1].6) LES(TIT_101_Vessel_Temperature,Vessel_Low_Low_Temperature_Setpoint) ,XIC(Vessel_2_Selected) XIO(Alarms[1].19) LES(TIT_201_Vessel_Temperature,Vessel_Low_Low_Temperature_Setpoint) ,XIC(Vessel_3_Selected) XIO(Alarms[1].20) LES(TIT_301_Vessel_Temperature,Vessel_Low_Low_Temperature_Setpoint) ]OTL(Alarms[1].11);
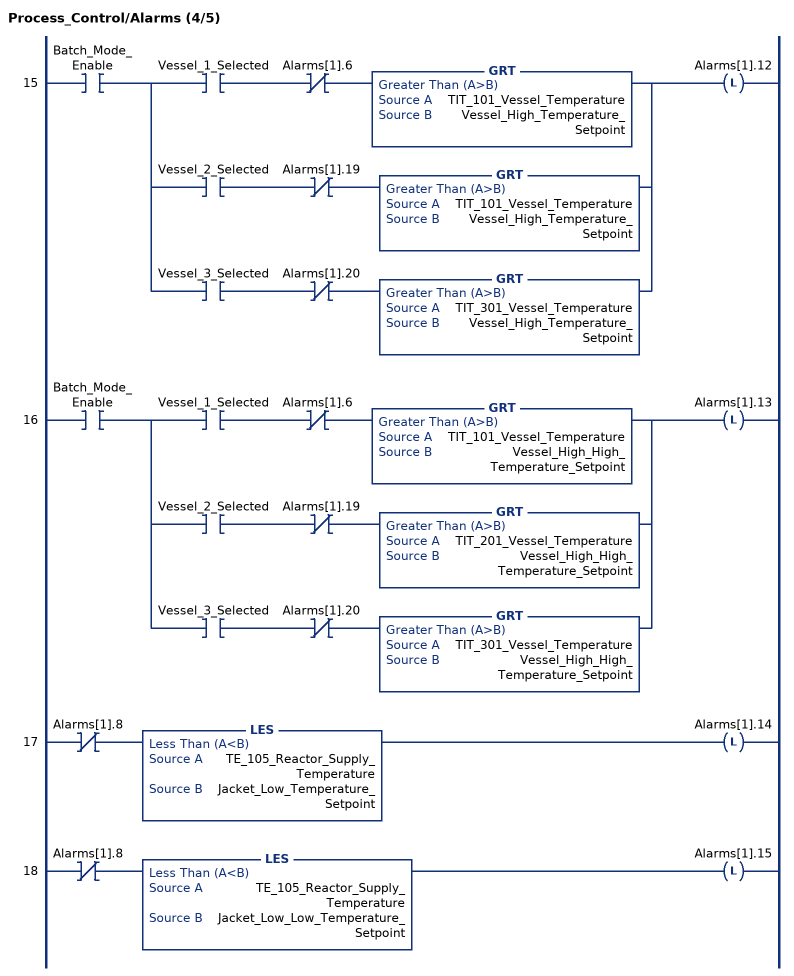
   15: XIC(Batch_Mode_Enable)[XIC(Vessel_1_Selected) XIO(Alarms[1].6) GRT(TIT_101_Vessel_Temperature,Vessel_High_Temperature_Setpoint) ,XIC(Vessel_2_Selected) XIO(Alarms[1].19) GRT(TIT_101_Vessel_Temperature,Vessel_High_Temperature_Setpoint) ,XIC(Vessel_3_Selected) XIO(Alarms[1].20) GRT(TIT_301_Vessel_Temperature,Vessel_High_Temperature_Setpoint) ]OTL(Alarms[1].12);
   16: XIC(Batch_Mode_Enable)[XIC(Vessel_1_Selected) XIO(Alarms[1].6) GRT(TIT_101_Vessel_Temperature,Vessel_High_High_Temperature_Setpoint) ,XIC(Vessel_2_Selected) XIO(Alarms[1].19) GRT(TIT_201_Vessel_Temperature,Vessel_High_High_Temperature_Setpoint) ,XIC(Vessel_3_Selected) XIO(Alarms[1].20) GRT(TIT_301_Vessel_Temperature,Vessel_High_High_Temperature_Setpoint) ]OTL(Alarms[1].13);
   17: XIO(Alarms[1].8)LES(TE_105_Reactor_Supply_Temperature,Jacket_Low_Temperature_Setpoint)OTL(Alarms[1].14);
   18: XIO(Alarms[1].8)LES(TE_105_Reactor_Supply_Temperature,Jacket_Low_Low_Temperature_Setpoint)OTL(Alarms[1].15);
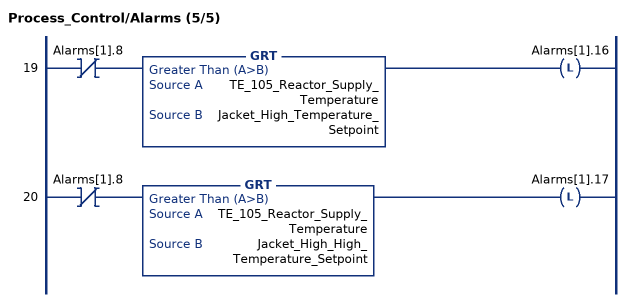
   19: XIO(Alarms[1].8)GRT(TE_105_Reactor_Supply_Temperature,Jacket_High_Temperature_Setpoint)OTL(Alarms[1].16);
   20: XIO(Alarms[1].8)GRT(TE_105_Reactor_Supply_Temperature,Jacket_High_High_Temperature_Setpoint)OTL(Alarms[1].17);
END_ROUTINE

ROUTINE Config   (* ladder *)
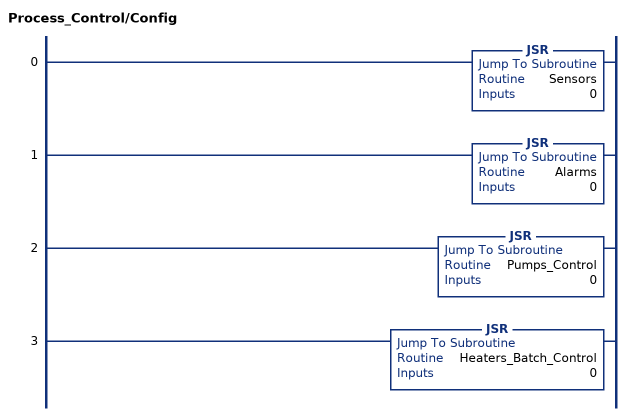
   0: JSR(Sensors,0);
   1: JSR(Alarms,0);
   2: JSR(Pumps_Control,0);
   3: JSR(Heaters_Batch_Control,0);
END_ROUTINE
